// TIA Portal V21 export
DATA_BLOCK "IDB_AnaUnused"   // DB13
// stored: InstanceOfName FB_AnaUnused, InstanceOfType FB
"FB_AnaUnused"
   // VAR_INPUT
   //    UsedInput : Int;
   //    UnusedInput : Int;
   // END_VAR
   // VAR_OUTPUT
   //    Result : Int;
   // END_VAR
   // VAR
   //    UnusedStatic : Int;
   // END_VAR
BEGIN
END_DATA_BLOCK
